(* IEC 61131-3 sources: ZPLC/packages/zplc-ide/projects/tank_level_starter/src, 1 file *)

(* ---- TankLevel.st ---- *)
PROGRAM TankLevel
VAR_INPUT AutoEnable AT %I0.0 : BOOL; LevelLow AT %I0.1 : BOOL; LevelHigh AT %I0.2 : BOOL; PumpFault AT %I0.3 : BOOL; EStop AT %I0.4 : BOOL; Reset AT %I0.5 : BOOL; END_VAR
VAR_OUTPUT Pump AT %Q0.0 : BOOL; Alarm AT %Q0.1 : BOOL; END_VAR
(* Exercise: keep the pump running from LevelLow until LevelHigh, latch Alarm on PumpFault or EStop, and release it only with a Reset pressed after the fault input has cleared. *)
Pump := AutoEnable AND LevelLow;
Alarm := FALSE;
END_PROGRAM
